(* IEC 61131-3 sources: llm-plc-st-eval/data/definitivo/gemini-3.1-pro-preview/C4/zero_shot, 3 files *)

(* ---- ejec_1.st ---- *)
### Descripción del Bloque de Función

El bloque de función `FB_D` es un **controlador de alternancia y respaldo (Duty/Standby o Lead/Lag) para un sistema redundante de dos bombas**. Su función principal es distribuir el desgaste de los equipos alternando la bomba principal (bomba de turno) cada vez que se recibe una nueva señal de `demanda`. Además, incorpora una lógica de alta disponibilidad (failover): si la bomba a la que le corresponde operar presenta una falla, el bloque arranca automáticamente la bomba de respaldo (siempre y cuando esta no esté en falla también) y activa una alarma. Esta lógica es ideal para aplicaciones industriales críticas como sistemas de bombeo de agua potable, cárcamos de rebombeo, circuitos de refrigeración (HVAC) o sistemas de lubricación, donde se requiere asegurar el suministro continuo y equilibrar las horas de uso de los motores.

---

### Código Estructurado (ST) Comentado

```iecst
// Bloque de función para alternancia y respaldo de dos bombas
FUNCTION_BLOCK FB_D
VAR_INPUT
    demanda : BOOL; // Señal de petición de arranque del sistema (ej. presostato, nivel, etc.)
    falla1 : BOOL;  // Señal de falla de la bomba 1 (ej. guardamotor, térmico)
    falla2 : BOOL;  // Señal de falla de la bomba 2 (ej. guardamotor, térmico)
END_VAR
VAR_OUTPUT
    bomba1 : BOOL;   // Comando de arranque para la bomba 1
    bomba2 : BOOL;   // Comando de arranque para la bomba 2
    almFalla : BOOL; // Indicador de alarma (se activa si la bomba en turno falla)
END_VAR
VAR
    turno : BOOL;    // Memoria interna para alternar el turno (FALSE = Bomba 2, TRUE = Bomba 1)
    fDem : R_TRIG;   // Detector de flanco de subida para la señal de demanda
END_VAR

// 1. Detección del flanco de subida de la demanda
fDem(CLK := demanda);

// 2. Lógica de alternancia
// Cada vez que entra una nueva demanda, se invierte el turno para equilibrar el desgaste
IF fDem.Q THEN
    turno := NOT turno;
END_IF

// 3. Lógica de control de bombas y respaldo (Failover)
IF demanda THEN

    // Si hay demanda, evaluamos de quién es el turno
    IF turno THEN
        // TURNO DE LA BOMBA 1
        // La bomba 1 arranca si no tiene falla
        bomba1 := NOT falla1;
        // La bomba 2 entra al quite (respaldo) si la bomba 1 falla y la bomba 2 está sana
        bomba2 := falla1 AND NOT falla2;
        // Se activa la alarma si la bomba titular (bomba 1) presenta falla
        almFalla := falla1;

    ELSE
        // TURNO DE LA BOMBA 2
        // La bomba 2 arranca si no tiene falla
        bomba2 := NOT falla2;
        // La bomba 1 entra al quite (respaldo) si la bomba 2 falla y la bomba 1 está sana
        bomba1 := falla2 AND NOT falla1;
        // Se activa la alarma si la bomba titular (bomba 2) presenta falla
        almFalla := falla2;
    END_IF

ELSE
    // 4. Estado de reposo
    // Si no hay demanda, se apagan ambas bombas y se limpia la alarma de turno
    bomba1 := FALSE;
    bomba2 := FALSE;
    almFalla := FALSE;
END_IF

END_FUNCTION_BLOCK
```

(* ---- ejec_2.st ---- *)
### Descripción del Bloque de Función

El bloque de función `FB_D` implementa un sistema de control de alternancia y respaldo automático (configuración *duty/standby*) para un sistema de dos bombas. Su función principal es alternar la bomba de trabajo cada vez que se recibe una nueva señal de demanda, lo que garantiza un desgaste mecánico uniforme entre ambos equipos a lo largo del tiempo. Además, incorpora una lógica de redundancia o "relevo" por falla: si la bomba a la que le corresponde operar presenta una avería, el sistema arranca automáticamente la bomba de respaldo (siempre y cuando esta no esté fallada también) y emite una señal de alarma. Esta lógica es ideal para aplicaciones industriales y comerciales de alta disponibilidad, tales como estaciones de bombeo de agua potable, cárcamos de rebombeo o achique, y circuitos de recirculación de agua helada o caliente en sistemas HVAC.

---

### Código Estructurado (Structured Text) Comentado

```iecst
(* Bloque de función para alternancia y respaldo de 2 bombas *)
FUNCTION_BLOCK FB_D
VAR_INPUT
    demanda : BOOL; // Señal de petición de arranque del sistema
    falla1  : BOOL; // Señal de avería/falla de la bomba 1
    falla2  : BOOL; // Señal de avería/falla de la bomba 2
END_VAR
VAR_OUTPUT
    bomba1   : BOOL; // Comando de arranque para la bomba 1
    bomba2   : BOOL; // Comando de arranque para la bomba 2
    almFalla : BOOL; // Alarma activa si la bomba en turno presenta falla
END_VAR
VAR
    turno : BOOL;   // Memoria para alternar el turno (FALSE = Bomba 2, TRUE = Bomba 1)
    fDem  : R_TRIG; // Detector de flanco de subida para la señal de demanda
END_VAR

// 1. Detección de nueva demanda para la alternancia
fDem(CLK := demanda); // Evalúa si la demanda pasó de FALSE a TRUE

// 2. Lógica de alternancia de turno
IF fDem.Q THEN
    turno := NOT turno; // Invierte el turno cada vez que inicia una nueva demanda
END_IF

// 3. Lógica de control de operación y respaldo
IF demanda THEN

    IF turno THEN
        // --- TURNO DE LA BOMBA 1 ---
        // La bomba 1 arranca si no tiene falla
        bomba1 := NOT falla1;
        // La bomba 2 entra como respaldo si la bomba 1 falla (y la 2 está sana)
        bomba2 := falla1 AND NOT falla2;
        // Se activa la alarma si la bomba titular (bomba 1) falló
        almFalla := falla1;

    ELSE
        // --- TURNO DE LA BOMBA 2 ---
        // La bomba 2 arranca si no tiene falla
        bomba2 := NOT falla2;
        // La bomba 1 entra como respaldo si la bomba 2 falla (y la 1 está sana)
        bomba1 := falla2 AND NOT falla1;
        // Se activa la alarma si la bomba titular (bomba 2) falló
        almFalla := falla2;
    END_IF

ELSE
    // 4. Condición de reposo (Sin demanda)
    // Se apagan ambas bombas y se limpia la alarma de falla de turno
    bomba1 := FALSE;
    bomba2 := FALSE;
    almFalla := FALSE;
END_IF

END_FUNCTION_BLOCK
```

(* ---- ejec_3.st ---- *)
### Descripción del Bloque de Función

El bloque de función `FB_D` implementa un sistema de control de **alternancia y respaldo (failover)** para un arreglo de dos bombas o motores. Su función principal es distribuir el desgaste de los equipos alternando la bomba "líder" (principal) cada vez que se detecta una nueva petición de arranque (flanco de subida en la señal de `demanda`). Además, cuenta con una lógica de redundancia de alta disponibilidad: si la bomba a la que le corresponde operar presenta una falla, el bloque arranca automáticamente la bomba de respaldo y activa una señal de alarma. Esta lógica es ideal para aplicaciones industriales como estaciones de bombeo de agua, sistemas de achique (cárcamos), compresores de aire o sistemas de refrigeración HVAC, donde se requiere asegurar el suministro continuo del proceso y prolongar la vida útil de los actuadores mediante un uso equilibrado.

---

### Código Comentado

```iecst
FUNCTION_BLOCK FB_D
VAR_INPUT
    demanda : BOOL; // Señal de petición de arranque (ej. presostato, interruptor de nivel, comando remoto)
    falla1 : BOOL;  // Señal de falla térmica o eléctrica de la bomba 1 (TRUE = en falla)
    falla2 : BOOL;  // Señal de falla térmica o eléctrica de la bomba 2 (TRUE = en falla)
END_VAR
VAR_OUTPUT
    bomba1 : BOOL;   // Comando de salida para energizar el contactor/variador de la bomba 1
    bomba2 : BOOL;   // Comando de salida para energizar el contactor/variador de la bomba 2
    almFalla : BOOL; // Señal de alarma que indica que la bomba líder actual ha fallado
END_VAR
VAR
    turno : BOOL;    // Memoria interna para alternar el turno (TRUE = turno bomba 1, FALSE = turno bomba 2)
    fDem : R_TRIG;   // Instancia del bloque detector de flanco de subida (Rising Trigger)
END_VAR

// 1. Detección de flanco de subida en la señal de demanda
fDem(CLK := demanda);

// 2. Lógica de alternancia (Flip-Flop)
// Cada vez que entra una nueva demanda, se invierte el turno para equilibrar el desgaste
IF fDem.Q THEN
    turno := NOT turno;
END_IF

// 3. Lógica principal de control y respaldo (Failover)
IF demanda THEN
    // Si hay demanda activa, evaluamos a quién le toca operar
    IF turno THEN
        // --- TURNO DE LA BOMBA 1 COMO LÍDER ---
        // La bomba 1 arranca si no tiene falla
        bomba1 := NOT falla1;
        // Si la bomba 1 falla, la bomba 2 entra como respaldo (siempre y cuando la 2 no esté en falla)
        bomba2 := falla1 AND NOT falla2;
        // Se activa la alarma si la bomba líder de este turno (bomba 1) presenta falla
        almFalla := falla1;
    ELSE
        // --- TURNO DE LA BOMBA 2 COMO LÍDER ---
        // La bomba 2 arranca si no tiene falla
        bomba2 := NOT falla2;
        // Si la bomba 2 falla, la bomba 1 entra como respaldo (siempre y cuando la 1 no esté en falla)
        bomba1 := falla2 AND NOT falla1;
        // Se activa la alarma si la bomba líder de este turno (bomba 2) presenta falla
        almFalla := falla2;
    END_IF
ELSE
    // 4. Estado de reposo
    // Si no hay demanda, se apagan ambas bombas y se limpia la alarma de falla de turno
    bomba1 := FALSE;
    bomba2 := FALSE;
    almFalla := FALSE;
END_IF
END_FUNCTION_BLOCK
```
